(*
SPDX-FileCopyrightText: c 2026 Oleksandr Tiutyk <trofimich@gmail.com>
SPDX-License-Identifier: MIT
License: https://opensource.org/license/mit
*)

(*!
<summary>Checks the concrete assignment failures and recovery with a matching buffer.</summary>
<description>
Uses one task and stays at a stable address while assertions are bound to this instance.
</description>
*)

{attribute 'no_assign'}
{attribute 'no_explicit_call' := 'do not call this function block directly'}
FUNCTION_BLOCK StringBuilderAssignmentFailureTest EXTENDS TOF_Testing.SingleCycleTest
VAR_STAT
	{attribute 'hide'}
	_ClassName : STRING := __POUNAME();
END_VAR
VAR
	_Builder : TOF_Core.StringBuilder;
END_VAR

(*!
<summary>Checks the concrete assignment failures and recovery with a matching buffer.</summary>
<description>
The builder is persistent so teardown can release its buffer after an unexpected hook exception.
</description>
*)
METHOD PROTECTED ExecuteTest
VAR
	wideTarget : WSTRING := "wide sentinel";
	shortTarget : STRING(10) := 'keep';
	exactTarget : STRING(16);

	exceptionCode : __SYSTEM.ExceptionCode;
	caught : TOF_Core.IException;
	typeException : TOF_Core.IArgumentTypeClassNotSupportedException;
	capacityException : TOF_Core.ITargetVariableMemoryOverflowException;
	copied : BOOL;
END_VAR
_Builder.AppendString255(value := 'String1234567890');

// Invoke a wrong-width target and check that the argument is rejected before modification.
__TRY
	_Builder.AssignToString(targetString := wideTarget);
__CATCH(exceptionCode)
	caught := TOF_Core.ExceptionManager.GetLastException(
		exceptionCode := exceptionCode,
		catchPointNamespaceName := NamespaceName,
		catchPointPOUName := __POUNAME(),
		catchPointPosition := __POSITION()
	);
__ENDTRY

Assert.ThatBool(
	actual := __QUERYINTERFACE(caught, typeException),
	message := "AssignToString must report an incompatible WSTRING target"
).IsTrue();
Assert.ThatBool(
	actual := wideTarget = "wide sentinel",
	message := "Wrong-width assignment must preserve the target"
).IsTrue();

caught := 0;

// Invoke an undersized STRING target and capture the documented capacity exception.
__TRY
	_Builder.AssignToString(targetString := shortTarget);
__CATCH(exceptionCode)
	caught := TOF_Core.ExceptionManager.GetLastException(
		exceptionCode := exceptionCode,
		catchPointNamespaceName := NamespaceName,
		catchPointPOUName := __POUNAME(),
		catchPointPosition := __POSITION()
	);
__ENDTRY

Assert.ThatBool(
	actual := __QUERYINTERFACE(caught, capacityException),
	message := "AssignToString must report insufficient capacity"
).IsTrue();
Assert.ThatBool(
	actual := shortTarget = 'keep',
	message := "Capacity rejection must preserve the target"
).IsTrue();

copied := _Builder.AssignToString(targetString := exactTarget);
Assert.ThatBool(
	actual := copied AND_THEN exactTarget = 'String1234567890',
	message := "The same builder must still copy successfully into the exact-fit target"
).IsTrue();
END_METHOD

(*!
<summary>Releases the builder buffer before reporting the case result.</summary>
<description>
Safe after partial initialization and after explicit cleanup in the scenario.
</description>
*)
METHOD PROTECTED AfterTest
_Builder.Clear(releaseMemory := TRUE);
END_METHOD

//! <summary>Borrows the concrete class name. Callers must not modify it.</summary>
{attribute 'monitoring' := 'call'}
PROPERTY ClassName : REFERENCE TO STRING
GET
ClassName REF= _ClassName;
END_GET
END_PROPERTY

//! <summary>Borrows the compiler-initialized namespace name. Callers must not modify it.</summary>
{attribute 'monitoring' := 'call'}
PROPERTY NamespaceName : REFERENCE TO STRING
GET
NamespaceName REF= CurrentNamespace.Name;
END_GET
END_PROPERTY

//! <summary>Reports the concrete instance size in bytes.</summary>
{attribute 'monitoring' := 'call'}
PROPERTY SelfSize : ULINT
GET
SelfSize := XSIZEOF(THIS^);
END_GET
END_PROPERTY

END_FUNCTION_BLOCK

(* stored: Version 1.1.0.1
   POU StringBuilderAssignmentFailureTest: Id {af43afb1-fb29-4628-80bd-e33350ddbf86}, SpecialFunc None
   Method ExecuteTest: Id {9586f9ed-636c-42d3-ade8-c23ea2a757d3}
   Method AfterTest: Id {419d7ab1-93fe-4a83-a3b0-5d6f3701210c}
   Property ClassName: Id {09da30b5-3f15-4e23-a65e-8e2abc3e1862}
   Get Get: Id {adf34ab2-3134-4b20-b629-f19a70459d39}
   Property NamespaceName: Id {450f895f-49ba-4a18-9226-05873ea58001}
   Get Get: Id {ab4d2755-e6a3-4b1b-85a0-a4da2a1d67ce}
   Property SelfSize: Id {d5a2d51e-a138-4338-a97c-811d76fed423}
   Get Get: Id {8372e739-a2ea-4f77-8a20-a90793849d7d} *)
